(*
SPDX-FileCopyrightText: c 2026 Oleksandr Tiutyk <trofimich@gmail.com>
SPDX-License-Identifier: MIT
License: https://opensource.org/license/mit
*)

(*!
<summary>Checks FIFO head, copy independence, length and capacity during dynamic growth.</summary>
<description>
Owns a dynamic queue and copied payloads at a stable address. Run from one task.
Teardown clears surviving entries and releases dynamic capacity.
</description>
*)

{attribute 'no_assign'}
{attribute 'no_explicit_call' := 'do not call this function block directly'}
FUNCTION_BLOCK DynamicQueueEnqueueAndPeekTest EXTENDS TOF_Testing.SingleCycleTest
VAR_STAT
	{attribute 'hide'}
	_ClassName : STRING := __POUNAME();
END_VAR
VAR
	_Queue : TOF_Collections.Queue<0>(valueValidator := 0);
END_VAR

(*!
<summary>Checks FIFO head, copy independence, length and capacity during dynamic growth.</summary>
*)
METHOD PROTECTED ExecuteTest
VAR
	values : ARRAY [1..4] OF INT := [11, 22, 33, 44];
END_VAR
_Queue.DefaultDynamicAllocationElementCount := BYTE#2;

_Queue.EnqueueCopy(value := values[1]);
values[1] := 111;

Assert.ThatInt(
	actual := _Queue.Peek().AsInt(),
	message := "Changing the source must preserve the copied head"
).ToBe(expected := INT#11);

Assert.ThatDInt(
	actual := _Queue.Capacity,
	message := "First enqueue must allocate two slots"
).ToBe(expected := DINT#2);

_Queue.EnqueueCopy(value := values[2]);

Assert.ThatInt(
	actual := _Queue.Peek().AsInt(),
	message := "Second enqueue must preserve the head"
).ToBe(expected := INT#11);

Assert.ThatBool(
	actual := _Queue.Full,
	message := "A dynamic queue must report not full when length equals capacity"
).IsFalse();

_Queue.EnqueueCopy(value := values[3]);

Assert.ThatInt(
	actual := _Queue.Peek().AsInt(),
	message := "Growing the descriptor buffer must preserve the head"
).ToBe(expected := INT#11);

Assert.ThatDInt(
	actual := _Queue.Length,
	message := "Three enqueues must produce three entries"
).ToBe(expected := DINT#3);

Assert.ThatDInt(
	actual := _Queue.Capacity,
	message := "Third enqueue must grow to four slots"
).ToBe(expected := DINT#4);

Assert.ThatInt(
	actual := _Queue.GetByIndex(index := 2).AsInt(),
	message := "Third enqueue must append the tail"
).ToBe(expected := values[3]);
END_METHOD

(*!
<summary>Clears the fixture before the runner publishes the result.</summary>
<description>
Also runs after an unexpected exception interrupts the case.
</description>
*)
METHOD PROTECTED AfterTest
_Queue.Clear();
END_METHOD

//! <summary>Borrows the concrete class name. Callers must not modify it.</summary>
{attribute 'monitoring' := 'call'}
PROPERTY ClassName : REFERENCE TO STRING
GET
ClassName REF= _ClassName;
END_GET
END_PROPERTY

//! <summary>Borrows the compiler-initialized namespace name. Callers must not modify it.</summary>
{attribute 'monitoring' := 'call'}
PROPERTY NamespaceName : REFERENCE TO STRING
GET
NamespaceName REF= CurrentNamespace.Name;
END_GET
END_PROPERTY

//! <summary>Reports the concrete instance size in bytes.</summary>
{attribute 'monitoring' := 'call'}
PROPERTY SelfSize : ULINT
GET
SelfSize := XSIZEOF(THIS^);
END_GET
END_PROPERTY

END_FUNCTION_BLOCK

(* stored: Version 1.1.0.1
   POU DynamicQueueEnqueueAndPeekTest: Id {a0217c3b-0bdc-413f-ae83-eb1b3ef51786}, SpecialFunc None
   Method ExecuteTest: Id {14841a3b-fe19-4f72-b4f9-ffc04d0ee69f}
   Method AfterTest: Id {b0e9403f-3ead-4bde-bf0d-4a7c24fad920}
   Property ClassName: Id {868ede50-aafa-4496-9b30-8d04a9d0713d}
   Get Get: Id {30492c36-7025-42dd-b0fc-0ed8e20426bc}
   Property NamespaceName: Id {09adc502-8e5c-466e-a379-79f5cfe77ff5}
   Get Get: Id {5e09480d-b4a4-4652-90f7-c403dd41b053}
   Property SelfSize: Id {1a8a9ce2-9303-4de7-80d7-88661c1c24eb}
   Get Get: Id {fca45f5c-c78f-4919-8b23-1d289f303330} *)
